PROGRAM main
  VAR
    B1 AT %IX0.0   : BOOL; (* sensor de cajas *)
    KM1 AT %QX0.0  : BOOL; (* banda (bobina 00001 para la PC) *)
    CAJAS AT %MW0  : INT; (* holding 40001: cajas contadas *)
    MARCHA AT %MW1 : INT; (* holding 40002: marcha, la escribe la PC *)
    META AT %MW2   : INT; (* holding 40003: meta de cajas, la escribe la PC *)
    F_CAJA         : R_TRIG;
    HAY_META       : BOOL; (* la PC fijó una meta *)
    LLENO          : BOOL; (* se llegó a la meta *)
  END_VAR
  VAR  (* added by the conversion: wires and edge detectors of the diagram *)
    R_TRIG1 : R_TRIG;
  END_VAR

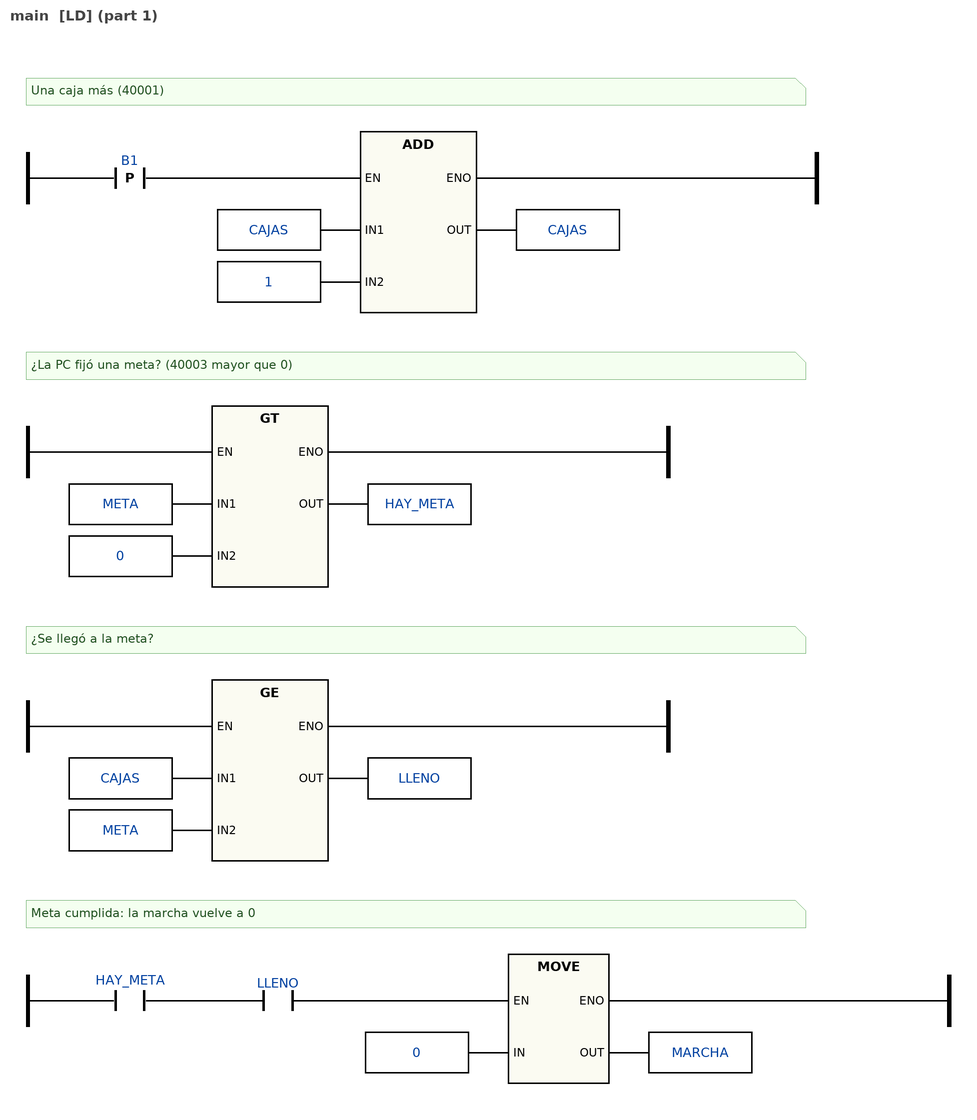
(* LD diagram, written out as Structured Text *)
(* Una caja más (40001) *)
R_TRIG1(CLK := B1);
IF R_TRIG1.Q THEN CAJAS := CAJAS + 1; END_IF;
(* ¿La PC fijó una meta? (40003 mayor que 0) *)
HAY_META := META > 0;
(* ¿Se llegó a la meta? *)
LLENO := CAJAS >= META;
(* Meta cumplida: la marcha vuelve a 0 *)
IF HAY_META AND LLENO THEN MARCHA := 0; END_IF;
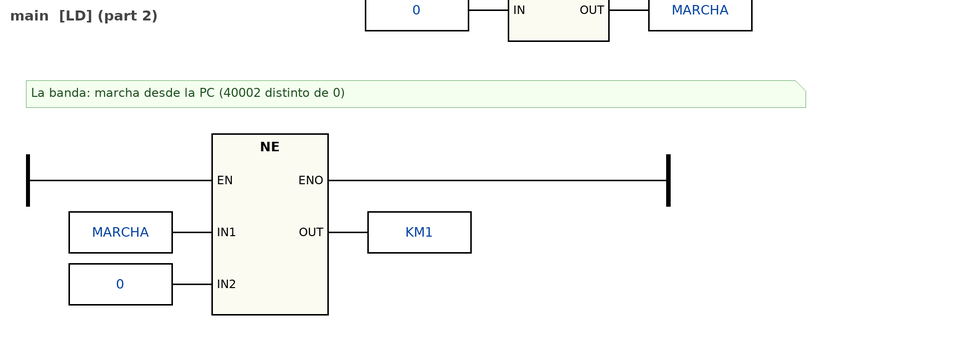
(* La banda: marcha desde la PC (40002 distinto de 0) *)
KM1 := MARCHA <> 0;
END_PROGRAM
